// TwinCAT 3 PLC project PLC1
// ProgramVersion: 3.1.4024.0
// libraries:
//   Tc2_MC2, * (Beckhoff Automation GmbH)
//   Tc2_Standard, * (Beckhoff Automation GmbH)
//   Tc2_System, * (Beckhoff Automation GmbH)
//   Tc2_TcpIp, * (Beckhoff Automation GmbH)
//   Tc3_Module, * (Beckhoff Automation GmbH)
// project tree:
//   DUTs/ E_MelsecDevice.TcDUT, ST_MelsecSession.TcDUT, ST_Point2D.TcDUT, ST_QD75_Command.TcDUT, ST_QD75_Feedback.TcDUT
//   GVLs/ GVL.TcGVL
//   / PlcTask.TcTTO
//   POUs/ FB_ConveyorEncoder.TcPOU, FB_ConveyorTracking4Pt.TcPOU, FB_EziServoControl.TcPOU, FB_MelsecRead.TcPOU, FB_MelsecTcpConfig.TcPOU, FB_MelsecWrite.TcPOU, FB_QD75CommandPublisher.TcPOU, MAIN.TcPOU
// real-time tasks:
//   TASK PlcTask: cycle T#10ms, priority 20, ADS port 350
// motion (NC):
//   TASK NC-Task 1 SAF: cycle T#2ms, priority 4, ADS port 501
//   TASK NC-Task 1 SVB: cycle T#10ms, priority 8, ADS port 511
//   AXIS Axis 1 (id 2)
//     General: UnitName=Degree
//     Velo: Maximum=50000
//     OtherSettings: AllowMotionCmdToSlave=true
//     encoder EncType=19
//       EncPara: ScaleFactorNumerator=360, ScaleFactorDenominator=10000, MaxCount=#xffffffff
//     drive DrvType=16
//       DrvPara: MaxCount=#xffffffff, DriveControlDWord=#x00020000
//         Analog: VeloReferenz=60000, TorqueSetpointScale=10, ScaleFactorActTorque=0.1
//         TimeComp: TaskDelayCycles=1
//     controller CtrType=1
//       CtrPara: PriorControlFactor=1
//         PosDiffControl: Range=60, Time=0.05
//         Observer: BandWidth=20
// I/O:
//   DEVICE Device 2 (EtherCAT), AmsNetId 10.81.27.140.3.1
//     Box 1 (NA-9286,Crevis) [NA-9286 EtherCAT Adapter, Crevis]
//       modules: Module 1 (ST-5101), Module 2 (ST-1228), Module 3 (ST-1228), Module 4 (ST-1228), Module 5 (ST-1228), Module 6 (ST-1228), Module 7 (ST-2318), Module 8 (ST-2318), Module 9 (ST-2318), Module 10 (ST-2318), Module 11 (ST-4424), Module 12 (ST-5114), Module 13 (ST-3214)
//     Drive 2 (Ezi-SERVO2 EtherCAT) [Ezi-SERVO2 EtherCAT]
// variable links:
//   NC-Task 1 SAF/Axes/Axis 1 <-> Device 2 (EtherCAT)/Drive 2 (Ezi-SERVO2 EtherCAT)
//     Drive/Inputs/In/nDcOutputTime <-> InfoData/DcOutputShift
//     Drive/Inputs/In/nState1 <-> CSP Inputs/Status Word
//     Drive/Inputs/In/nState2 <-> CSP Inputs/Status Word @bit 8
//     Drive/Inputs/In/nState4 @bit 1 <-> WcState/InputToggle
//     Drive/Inputs/In/nState4 <-> WcState/WcState
//     Drive/Outputs/Out/nCtrl1 <-> CSP Outputs/Control Word
//     Drive/Outputs/Out/nCtrl2 <-> CSP Outputs/Control Word @bit 8
//     Drive/Outputs/Out/nDataOut1 <-> CSP Outputs/Target Position
//     Enc/Inputs/In/nDataIn1 <-> CSP Inputs/Position Actual Value
//     Enc/Inputs/In/nDataIn3 <-> CSP Inputs/Touch probe 1 positive value
//     Enc/Inputs/In/nDataIn5 <-> CSP Inputs/Touch probe 2 positive value
//     Enc/Inputs/In/nDcInputTime <-> InfoData/DcInputShift
//     Enc/Inputs/In/nState4 @bit 1 <-> WcState/InputToggle
//     Enc/Inputs/In/nState4 <-> WcState/WcState
//     Enc/Inputs/In/nState5 <-> CSP Inputs/Touch probe status
//     Enc/Inputs/In/nState6 <-> CSP Inputs/Touch probe status @bit 8
//     Enc/Outputs/Out/nCtrl5 <-> CSP Outputs/Touch probe function
//     Enc/Outputs/Out/nCtrl6 <-> CSP Outputs/Touch probe function @bit 8
//   PLC1/PLC1 Instance <-> Device 2 (EtherCAT)/Box 1 (NA-9286,Crevis)
//     PlcTask Inputs/GVL.aIn[{0..15}] <-> Module 12 (ST-5114)/Input(s)/Byte {0..15}  (16 links)
//     PlcTask Outputs/GVL.aOut[{0..3}] <-> Module 12 (ST-5114)/Output(s)/Byte {0..3}  (4 links)
//   PLC1/PLC1 Instance <-> NC-Task 1 SAF/Axes/Axis 1
//     PlcTask Inputs/MAIN.Axis1.NcToPlc <-> Outputs/ToPlc
//     PlcTask Outputs/MAIN.Axis1.PlcToNc <-> Inputs/FromPlc

CONFIGURATION PLC1
    RESOURCE PLC ON TwinCAT3
        TASK PlcTask(INTERVAL := T#10ms, PRIORITY := 20);
        PROGRAM MAIN WITH PlcTask : MAIN;
    END_RESOURCE
END_CONFIGURATION

// ---- DUTs/E_MelsecDevice.TcDUT
// Mã định danh vùng nhớ phần cứng Mitsubishi theo chuẩn MC Protocol Binary 3E Frame
TYPE E_MelsecDevice :
(
    DEV_D   := 16#A8, // Thanh ghi dữ liệu D (Data Register) - Word
    DEV_M   := 16#90, // Rơ-le nội bộ M (Internal Relay) - Bit / Word
    DEV_W   := 16#B4, // Thanh ghi liên kết W (Link Register) - Word
    DEV_R   := 16#AF, // Thanh ghi tệp R (File Register) - Word
    DEV_ZR  := 16#B0, // Thanh ghi tệp liên tục ZR (File Register Consecutive) - Word
    DEV_X   := 16#9C, // Ngõ vào vật lý X (Input) - Bit
    DEV_Y   := 16#9D, // Ngõ ra vật lý Y (Output) - Bit
    DEV_B   := 16#A0, // Rơ-le liên kết B (Link Relay) - Bit / Word
    DEV_L   := 16#92, // Rơ-le chốt L (Latch Relay) - Bit
    DEV_TN  := 16#C2, // Giá trị hiện tại Timer TN (Timer Current Value) - Word
    DEV_CN  := 16#C5  // Giá trị hiện tại Counter CN (Counter Current Value) - Word
);
END_TYPE

// ---- DUTs/ST_MelsecSession.TcDUT
TYPE ST_MelsecSession :
STRUCT
    hSocket     : T_HSOCKET; // Socket TCP dùng chung
    bConnected  : BOOL;      // TRUE khi đã kết nối PLC
    bBusy       : BOOL;      // TRUE khi Read hoặc Write đang giao dịch
    bError      : BOOL;      // Lỗi cuối cùng
    nErrorID    : UDINT;     // Mã lỗi cuối cùng
END_STRUCT
END_TYPE

// ---- DUTs/ST_Point2D.TcDUT
TYPE ST_Point2D :
STRUCT
    X : LREAL; // Tọa độ X (mm)
    Y : LREAL; // Tọa độ Y (mm)
END_STRUCT
END_TYPE

// ---- DUTs/ST_QD75_Command.TcDUT
TYPE ST_QD75_Command :
STRUCT
    Target_X       : DINT; // D100..D101: Tọa độ đón đầu trục X (0.1 um)
    Target_Y       : DINT; // D102..D103: Tọa độ trục Y đỉnh (0.1 um)
    Target_Z_Down  : DINT; // D104..D105: Độ cao hạ chấm keo (0.1 um, 4.0mm = 40000)
    Speed_Approach : DINT; // D106..D107: Vận tốc bay nội suy 3 trục (0.01 mm/min, 500mm/s = 3000000)
    Speed_Sync     : DINT; // D108..D109: Vận tốc đồng tốc trục X khi chấm keo (= V_conv * 6000)
    DeltaX_Sync    : DINT; // D110..D111: Quãng đường trượt đồng tốc 60ms (0.1 um)
    Target_Z_Safe  : DINT; // D112..D113: Độ cao an toàn khi rút kim (0.1 um, 0.0mm = 0)
    Vertex_Index   : INT;  // D114: Thứ tự đỉnh đang làm (1..4)
END_STRUCT
END_TYPE

// ---- DUTs/ST_QD75_Feedback.TcDUT
TYPE ST_QD75_Feedback :
STRUCT
    Ack_Done    : BOOL; // M1001: PLC-Q báo Point 3 hoàn tất
    Robot_Busy  : BOOL; // M102: PLC-Q đang kiểm tra/nạp/chạy
    In_Position : BOOL; // M103: Đỉnh đã hoàn tất, chờ Master hạ M1000
    Robot_Alarm : BOOL; // M104: QD75 hoặc kiểm tra biên báo lỗi
END_STRUCT
END_TYPE

// ---- GVLs/GVL.TcGVL
VAR_GLOBAL
    aIn  AT %I* : ARRAY[0..15] OF BYTE;  // TxPDO 16 byte
    aOut AT %Q* : ARRAY[0..3]  OF BYTE;  // RxPDO 4 byte
END_VAR

// ---- POUs/MAIN.TcPOU
PROGRAM MAIN
VAR
    // ================================================================
    // 1. KẾT NỐI TCP VỚI CPU MITSUBISHI Q06UDEH (CỔNG 5010)
    // ================================================================
    stMelsec            : ST_MelsecSession; // Session TCP dùng chung
    fbMelsecConfig      : FB_MelsecTcpConfig;

    bTcpEnable          : BOOL := TRUE;     // Tự động kết nối và duy trì kết nối mạng
    sPlcQ_IP            : STRING(15) := '192.168.3.39'; // IP của PLC-Q
    nPlcQ_Port          : UDINT := 5010;   // Cổng Port MC Protocol 5010

    bPlcQConnected      : BOOL;             // ĐÈN BÁO: TRUE = Đã thông mạng với PLC-Q
    bPlcQError          : BOOL;
    nPlcQErrorID        : UDINT;

    // ================================================================
    // 2. TEST TRUYỀN THÔNG THỦ CÔNG SANG PLC-Q (KHI bStartGlueCycle = FALSE)
    // ================================================================
    bTest_WriteD100     : BOOL := FALSE;    // Click đúp TRUE -> Ghi nTest_D100_Val vào D100-D101
    nTest_D100_Val      : DINT := 100;      // Số 32-bit gửi thử sang D100
    bTest_WriteM1000    : BOOL := FALSE;    // Click đúp TRUE -> Ghi bit M1000
    bTest_M1000_Val     : BOOL := TRUE;     // Giá trị bit M1000 muốn ghi (TRUE=ON, FALSE=OFF)
    bTest_ReadM1001     : BOOL := FALSE;    // Click đúp TRUE -> Đọc bit M1001 từ PLC-Q
    bTest_M1001_Result  : BOOL;             // Giá trị M1001 đọc được từ PLC-Q

    // ================================================================
    // 3. ENCODER BĂNG TẢI: ST-5114 MODULE 12
    // ================================================================
    fbConveyor          : FB_ConveyorEncoder;

    nEncoderPulse       : UINT;            // Số xung Encoder hiện tại
    nEncoderDelta       : INT;             // Xung thay đổi trong 10 ms
    rConveyorSpeed      : LREAL;           // Vận tốc băng tải lọc mượt, mm/s
    rConveyorSpeedMPM   : LREAL;           // Vận tốc băng tải, m/phút
    rConveyorDist       : LREAL;           // Tổng quãng đường băng tải, mm

    // ================================================================
    // 4. EZI-SERVO: TRỤC QUAY ĐƠN VỊ DEGREE
    // ================================================================
    Axis1               : AXIS_REF;

    fbServo             : FB_EziServoControl;

    bServo_Enable       : BOOL := TRUE;     // TRUE = Servo ON / giữ cốt
    bServo_Reset        : BOOL := FALSE;    // TRUE một chu kỳ = Reset Alarm
    bServo_JogFwd       : BOOL := FALSE;    // TRUE = chạy thuận
    bServo_JogBwd       : BOOL := FALSE;    // TRUE = chạy nghịch

    rServo_Speed        : LREAL := 100.0;   // Degree/s
    rServo_Acc          : LREAL := 400.0;   // Degree/s2
    rServo_Dec          : LREAL := 400.0;   // Degree/s2

    bServo_Ready        : BOOL;             // TRUE = Servo ON
    rServo_ActPos_Deg   : LREAL;            // Góc thực tế, Degree
    rServo_ActVel_Deg_s : LREAL;            // Vận tốc thực tế, Degree/s

    // ================================================================
    // 5. TRACKING 4 ĐIỂM: CAMERA + ENCODER
    // ================================================================
    fbTracking4Pt       : FB_ConveyorTracking4Pt;

    bSystemReset        : BOOL := FALSE;    // TRUE một chu kỳ: reset mốc phần mềm về 0
    // Camera giả lập test
    bCameraTrigger      : BOOL := FALSE;    // FALSE -> TRUE: chốt sản phẩm mới
    rCameraCenterX      : LREAL := 50.0;    // Tâm phôi X, mm
    rCameraCenterY      : LREAL := 85.0;    // Tâm phôi Y, mm
    rCameraAngleDeg     : LREAL := 0.0;     // Góc phôi, Degree
    rProductLength      : LREAL := 40.0;    // mm
    rProductWidth       : LREAL := 40.0;    // mm

    // Kết quả debug Tracking
    bProductValid       : BOOL;
    nPulseAtCamera      : UINT;
    nPulseTravel        : INT;
    rPartTravel_mm      : LREAL;

    aCornerBase         : ARRAY[1..4] OF ST_Point2D;
    aCornerNow          : ARRAY[1..4] OF ST_Point2D;

    // ================================================================
    // 6. QD75 COMMAND PUBLISHER: ĐIỀU PHỐI 4 ĐỈNH SANG PLC-Q
    // ================================================================
    fbPublisher         : FB_QD75CommandPublisher;

    // Lệnh chu trình chấm keo
    bStartGlueCycle     : BOOL := FALSE;   // FALSE -> TRUE: kích chạy chu trình 4 đỉnh
    bAbortGlueCycle     : BOOL := FALSE;   // TRUE: dừng khẩn cấp (ghi M105)

    // Trạng thái giám sát chu trình
    bGlueCycleBusy      : BOOL;            // Đang chạy 4 đỉnh
    bGlueCycleDone      : BOOL;            // Hoàn tất cả 4 đỉnh
    bGlueCycleError     : BOOL;            // Báo lỗi
    nGlueCurVertex      : INT;             // Đỉnh đang thực hiện (1..4)
    nGlueErrorCode      : INT;             // Mã lỗi (501..503, 900..921)
END_VAR

// ================================================================
// 1. TCP CONFIG: Kết nối / tự reconnect đến PLC-Q
// ================================================================
fbMelsecConfig(
    bEnable     := bTcpEnable,
    sRemoteHost := sPlcQ_IP,
    nRemotePort := nPlcQ_Port,
    stSession   := stMelsec
);

// Biến trạng thái đưa ra ngoài để Online debug dễ
bPlcQConnected := stMelsec.bConnected;
bPlcQError     := stMelsec.bError;
nPlcQErrorID   := stMelsec.nErrorID;


// ================================================================
// 2. ENCODER BĂNG TẢI: ST-5114 INPUT BYTE 0 + BYTE 1
// ================================================================
fbConveyor(
    bByte0          := GVL.aIn[0],
    bByte1          := GVL.aIn[1],
    rK_mm           := 0.476475,
    rCycleTime      := 0.01,

    nRawPulse       => nEncoderPulse,
    nDeltaPulse     => nEncoderDelta,
    rSpeed_mm_s     => rConveyorSpeed,
    rSpeed_m_min    => rConveyorSpeedMPM,
    rTotalDist_mm   => rConveyorDist
);


// ================================================================
// 3. EZI-SERVO: ENABLE, RESET, JOG VÀ GIÁM SÁT
// ================================================================
fbServo(
    Axis            := Axis1,
    bEnable         := bServo_Enable,
    bResetFault     := bServo_Reset,
    bJogFwd         := bServo_JogFwd,
    bJogBwd         := bServo_JogBwd,
    rTargetVelocity := rServo_Speed,
    rAcc            := rServo_Acc,
    rDec            := rServo_Dec,

    bReady          => bServo_Ready,
    rActPos_Deg     => rServo_ActPos_Deg,
    rActVel_Deg     => rServo_ActVel_Deg_s
);

IF bServo_Reset THEN
    bServo_Reset := FALSE;
END_IF;


// ================================================================
// 4. TRACKING 4 ĐIỂM: CAMERA + ENCODER
// ================================================================
fbTracking4Pt(
    bResetSystem   := bSystemReset,
    bCameraResult  := bCameraTrigger,
    rCenterX_mm    := rCameraCenterX,
    rCenterY_mm    := rCameraCenterY,
    rAngleDeg      := rCameraAngleDeg,
    rLength_mm     := rProductLength,
    rWidth_mm      := rProductWidth,

    nEncoderNow    := nEncoderPulse,
    rMmPerPulse    := 0.476475,
    rXMaxLimit_mm  := 180.0,

    bProductValid  => bProductValid,
    nPulseAtCamera => nPulseAtCamera,
    nPulseTravel   => nPulseTravel,
    rTravel_mm     => rPartTravel_mm,
    aCornerBase    => aCornerBase,
    aCornerNow     => aCornerNow
);

IF bSystemReset THEN
    bSystemReset := FALSE;
END_IF;


// ================================================================
// 5. QD75 COMMAND PUBLISHER: ĐIỀU PHỐI 4 ĐỈNH & TEST THỦ CÔNG
// ================================================================
fbPublisher(
    stSession           := stMelsec,
    bStartCycle         := bStartGlueCycle,
    bAbortCycle         := bAbortGlueCycle,

    // Tọa độ 4 góc thời gian thực từ khối Tracking
    aCornerNow          := aCornerNow,
    rConveyorSpeed_mm_s := rConveyorSpeed,

    // Động học
    rFlyTime_s          := 0.120,
    rApproachSpeed_mm_s := 500.0,
    rSyncTime_s         := 0.060,
    rZDown_mm           := 4.0,
    rZSafe_mm           := 0.0,

    // Chế độ test thủ công (chỉ có tác dụng khi bStartGlueCycle = FALSE)
    bManualWriteD100    := bTest_WriteD100,
    nD100_ManualVal     := nTest_D100_Val,
    bManualWriteM1000   := bTest_WriteM1000,
    bM1000_ManualVal    := bTest_M1000_Val,
    bManualReadM1001    := bTest_ReadM1001,

    // Giám sát
    bBusy               => bGlueCycleBusy,
    bDone               => bGlueCycleDone,
    bError              => bGlueCycleError,
    nErrorCode          => nGlueErrorCode,
    nCurrentVertex      => nGlueCurVertex,
    bM1001_ReadBack     => bTest_M1001_Result
);

// Tự động nhả cờ kích test sau khi lệnh được nhận
IF bTest_WriteD100 AND NOT fbPublisher.bManualWriteD100 THEN
    bTest_WriteD100 := FALSE;
END_IF;

IF bTest_WriteM1000 AND NOT fbPublisher.bManualWriteM1000 THEN
    bTest_WriteM1000 := FALSE;
END_IF;

IF bTest_ReadM1001 AND NOT fbPublisher.bManualReadM1001 THEN
    bTest_ReadM1001 := FALSE;
END_IF;

END_PROGRAM

// ---- POUs/FB_MelsecTcpConfig.TcPOU
FUNCTION_BLOCK FB_MelsecTcpConfig
VAR_INPUT
    bEnable         : BOOL := TRUE;                 // TRUE = duy trì kết nối
    sRemoteHost     : STRING(15) := '192.168.3.39'; // IP PLC-Q
    nRemotePort     : UDINT := 5010;               // Port MC Protocol
END_VAR
VAR_IN_OUT
    stSession       : ST_MelsecSession;             // Session TCP dùng chung
END_VAR
VAR
    fbConnect       : FB_SocketConnect;
    fbClose         : FB_SocketClose;
    tonRetry        : TON;

    nState          : INT := 0;
    bConnectError   : BOOL;
    nConnectErrorID : UDINT;
END_VAR

// State:
// 0 = chờ reconnect
// 1 = phát cạnh mở TCP
// 2 = chờ kết quả kết nối
// 10 = đã kết nối
// 20 = đóng socket khi Disable

CASE nState OF

    0: // Chờ 2 giây trước khi thử kết nối / kết nối lại
        stSession.bConnected := FALSE;
        stSession.bBusy      := FALSE;

        IF NOT bEnable THEN
            tonRetry(IN := FALSE);
            stSession.bError := FALSE;
        ELSE
            tonRetry(IN := TRUE, PT := T#2S);

            IF tonRetry.Q THEN
                tonRetry(IN := FALSE);
                stSession.bError   := FALSE;
                stSession.nErrorID := 0;
                nState := 1;
            END_IF
        END_IF


    1: // Cạnh lên mở TCP Socket
        fbConnect(
            sSrvNetId   := '',
            sRemoteHost := sRemoteHost,
            nRemotePort := nRemotePort,
            bExecute    := TRUE,
            tTimeout    := T#3S,
            bError      => bConnectError,
            nErrId      => nConnectErrorID,
            hSocket     => stSession.hSocket
        );

        stSession.bBusy := TRUE;
        nState := 2;


    2: // Chờ FB_SocketConnect hoàn thành
        fbConnect(
            sSrvNetId   := '',
            sRemoteHost := sRemoteHost,
            nRemotePort := nRemotePort,
            bExecute    := FALSE,
            tTimeout    := T#3S,
            bError      => bConnectError,
            nErrId      => nConnectErrorID,
            hSocket     => stSession.hSocket
        );

        IF NOT fbConnect.bBusy THEN
            stSession.bBusy := FALSE;

            IF bConnectError THEN
                stSession.bError   := TRUE;
                stSession.nErrorID := nConnectErrorID;
                stSession.hSocket.handle := 0;
                nState := 0; // Chờ 2 giây, tự thử lại
            ELSE
                stSession.bConnected := TRUE;
                stSession.bError     := FALSE;
                nState := 10;
            END_IF
        END_IF


    10: // TCP đang kết nối tốt
        stSession.bConnected := TRUE;

        IF NOT bEnable THEN
            nState := 20;
        END_IF


    20: // Đóng TCP Socket khi Disable
        fbClose(
            sSrvNetId := '',
            hSocket   := stSession.hSocket,
            bExecute  := TRUE,
            tTimeout  := T#3S
        );

        nState := 21;


    21: // Chờ đóng xong
        fbClose(
            sSrvNetId := '',
            hSocket   := stSession.hSocket,
            bExecute  := FALSE,
            tTimeout  := T#3S
        );

        IF NOT fbClose.bBusy THEN
            stSession.hSocket.handle := 0;
            stSession.bConnected     := FALSE;
            stSession.bBusy          := FALSE;
            nState := 0;
        END_IF

END_CASE

END_FUNCTION_BLOCK

// ---- POUs/FB_ConveyorEncoder.TcPOU
FUNCTION_BLOCK FB_ConveyorEncoder
VAR_INPUT
    bByte0          : BYTE;             // GVL.aIn[0]
    bByte1          : BYTE;             // GVL.aIn[1]
    rK_mm           : LREAL := 0.476475;// mm / xung (D=54.6mm, 360 xung)
    rCycleTime      : LREAL := 0.01;    // 10ms
END_VAR
VAR_OUTPUT
    nRawPulse       : UINT;             // Xung tức thời
    nDeltaPulse     : INT;              // Lệch xung mỗi 10ms
    rSpeed_mm_s     : LREAL;            // VẬN TỐC LỌC MƯỢT (mm/s)
    rSpeed_m_min    : LREAL;            // Vận tốc hiển thị (m/phút)
    rTotalDist_mm   : LREAL;            // TỔNG QUÃNG ĐƯỜNG (mm)
END_VAR
VAR
    nPrev           : UINT;
    bInit           : BOOL := TRUE;
    // Bộ lọc trượt 20 chu kỳ (200ms) để triệt tiêu hoàn toàn rung lắc
    aDeltaBuf       : ARRAY[0..19] OF INT;
    nBufIdx         : INT := 0;
    nSumDelta       : INT;
    nIdx            : INT;
    rSpeed_Avg_Raw  : LREAL;
END_VAR

// 1. Ghép 2 byte thành số xung 16-bit
nRawPulse := BYTE_TO_UINT(bByte1) * 256 + BYTE_TO_UINT(bByte0);

IF bInit THEN
    nPrev := nRawPulse;
    bInit := FALSE;
END_IF

// 2. Tính số xung lệch chu kỳ 10ms (chống tràn số)
nDeltaPulse := TO_INT(TO_DINT(nRawPulse) - TO_DINT(nPrev));
nPrev       := nRawPulse;

// 3. Bộ lọc trung bình trượt 20 chu kỳ (200ms)
aDeltaBuf[nBufIdx] := nDeltaPulse;
nBufIdx := (nBufIdx + 1) MOD 20;

nSumDelta := 0;
FOR nIdx := 0 TO 19 DO
    nSumDelta := nSumDelta + aDeltaBuf[nIdx];
END_FOR;

// 4. CẮT ZERO KHI DỪNG (DEAD-BAND):
// Nếu trong 200ms không có xung nào (băng tải dừng), ép thẳng về 0.0 ngay lập tức!
IF nSumDelta = 0 THEN
    rSpeed_mm_s  := 0.0;
    rSpeed_m_min := 0.0;
ELSE
    // Tính vận tốc trung bình trong 200ms
    rSpeed_Avg_Raw := (TO_LREAL(nSumDelta) * rK_mm) / 0.2;

    // Lọc mượt nhẹ
    rSpeed_mm_s    := rSpeed_mm_s + 0.2 * (rSpeed_Avg_Raw - rSpeed_mm_s);

    // LÀM TRÒN 1 CHỮ SỐ THẬP PHÂN (Để mắt nhìn thấy số đứng yên đầm chắc, ví dụ 100.2 mm/s)
    rSpeed_mm_s    := DINT_TO_LREAL(LREAL_TO_DINT(rSpeed_mm_s * 10.0)) / 10.0;
    rSpeed_m_min   := DINT_TO_LREAL(LREAL_TO_DINT((rSpeed_mm_s * 60.0 / 1000.0) * 10.0)) / 10.0;
END_IF;

// 5. Tổng quãng đường tích lũy (chuẩn xác 100% không lọc)
rTotalDist_mm := rTotalDist_mm + (TO_LREAL(nDeltaPulse) * rK_mm);

END_FUNCTION_BLOCK

// ---- POUs/FB_EziServoControl.TcPOU
FUNCTION_BLOCK FB_EziServoControl
VAR_INPUT
    bEnable         : BOOL := TRUE;
    bResetFault     : BOOL := FALSE;
    bJogFwd         : BOOL := FALSE;
    bJogBwd         : BOOL := FALSE;
    rTargetVelocity : LREAL := 100.0;
    rAcc            : LREAL := 400.0;
    rDec            : LREAL := 400.0;
END_VAR
VAR_IN_OUT
    Axis            : AXIS_REF;
END_VAR
VAR_OUTPUT
    bReady          : BOOL;
    rActPos_Deg     : LREAL;
    rActVel_Deg     : LREAL;
END_VAR
VAR
    fbPower         : MC_Power;
    fbMoveVelocity  : MC_MoveVelocity;
    fbHalt          : MC_Halt;
    fbReset         : MC_Reset;

    rTargetVel_Prev : LREAL;
    bVelChanged     : BOOL;
    fbTrigFwd       : R_TRIG;
    fbTrigBwd       : R_TRIG;
    fbTrigStop      : R_TRIG;
END_VAR

fbReset(Axis := Axis, Execute := bResetFault);

fbPower(
    Axis            := Axis,
    Enable          := bEnable,
    Enable_Positive := TRUE,
    Enable_Negative := TRUE,
    Override        := 100.0,
    Status          => bReady
);

fbTrigFwd(CLK := bJogFwd);
fbTrigBwd(CLK := bJogBwd);
fbTrigStop(CLK := (NOT bJogFwd AND NOT bJogBwd));

IF rTargetVelocity <> rTargetVel_Prev THEN
    bVelChanged     := TRUE;
    rTargetVel_Prev := rTargetVelocity;
ELSE
    bVelChanged     := FALSE;
END_IF

fbMoveVelocity(
    Axis         := Axis,
    Execute      := (fbTrigFwd.Q OR fbTrigBwd.Q OR (bVelChanged AND (bJogFwd OR bJogBwd))),
    Velocity     := rTargetVelocity,
    Acceleration := rAcc,
    Deceleration := rDec,
    Jerk         := 10000.0,
    Direction    := SEL(bJogBwd, MC_Positive_Direction, MC_Negative_Direction)
);

fbHalt(
    Axis         := Axis,
    Execute      := fbTrigStop.Q,
    Deceleration := rDec,
    Jerk         := 10000.0
);

rActPos_Deg := Axis.NcToPlc.ActPos;
rActVel_Deg := Axis.NcToPlc.ActVelo;

END_FUNCTION_BLOCK

// ---- POUs/FB_ConveyorTracking4Pt.TcPOU
FUNCTION_BLOCK FB_ConveyorTracking4Pt
VAR_INPUT
    bResetSystem     : BOOL;
    bCameraResult    : BOOL;
    rCenterX_mm      : LREAL;
    rCenterY_mm      : LREAL;
    rAngleDeg        : LREAL;
    rLength_mm       : LREAL := 40.0;
    rWidth_mm        : LREAL := 40.0;
    nEncoderNow      : UINT;
    rMmPerPulse      : LREAL := 0.476475;
    rXMaxLimit_mm    : LREAL := 180.0;
END_VAR

VAR_OUTPUT
    bProductValid    : BOOL;
    nPulseAtCamera   : UINT;
    nPulseTravel     : INT;
    rTravel_mm       : LREAL;
    aCornerBase      : ARRAY[1..4] OF ST_Point2D;
    aCornerNow       : ARRAY[1..4] OF ST_Point2D;
END_VAR

VAR
    fbCameraEdge     : R_TRIG;
    rRad             : LREAL;
    rCosA            : LREAL;
    rSinA            : LREAL;
    rHalfLength      : LREAL;
    rHalfWidth       : LREAL;
    nIndex           : INT;
    bFirstScan       : BOOL := TRUE;
END_VAR

// Reset mốc phần mềm một lần khi PLC khởi động hoặc khi bResetSystem kích.
IF bFirstScan OR bResetSystem THEN
    bFirstScan     := FALSE;
    bProductValid  := FALSE;
    nPulseAtCamera := nEncoderNow;
    nPulseTravel   := 0;
    rTravel_mm     := 0.0;

    FOR nIndex := 1 TO 4 DO
        aCornerBase[nIndex].X := 0.0;
        aCornerBase[nIndex].Y := 0.0;
        aCornerNow[nIndex].X  := 0.0;
        aCornerNow[nIndex].Y  := 0.0;
    END_FOR;
END_IF;

fbCameraEdge(CLK := bCameraResult);

// Camera chụp: chốt encoder và tính bốn góc gốc.
IF fbCameraEdge.Q THEN
    nPulseAtCamera := nEncoderNow;
    nPulseTravel   := 0;
    rTravel_mm     := 0.0;

    rRad   := rAngleDeg * 3.141592653589793 / 180.0;
    rCosA  := COS(rRad);
    rSinA  := SIN(rRad);
    rHalfLength := rLength_mm / 2.0;
    rHalfWidth  := rWidth_mm / 2.0;

    aCornerBase[1].X := rCenterX_mm + rHalfLength * rCosA - rHalfWidth * rSinA;
    aCornerBase[1].Y := rCenterY_mm + rHalfLength * rSinA + rHalfWidth * rCosA;
    aCornerBase[2].X := rCenterX_mm - rHalfLength * rCosA - rHalfWidth * rSinA;
    aCornerBase[2].Y := rCenterY_mm - rHalfLength * rSinA + rHalfWidth * rCosA;
    aCornerBase[3].X := rCenterX_mm - rHalfLength * rCosA + rHalfWidth * rSinA;
    aCornerBase[3].Y := rCenterY_mm - rHalfLength * rSinA - rHalfWidth * rCosA;
    aCornerBase[4].X := rCenterX_mm + rHalfLength * rCosA + rHalfWidth * rSinA;
    aCornerBase[4].Y := rCenterY_mm + rHalfLength * rSinA - rHalfWidth * rCosA;

    FOR nIndex := 1 TO 4 DO
        aCornerNow[nIndex] := aCornerBase[nIndex];
    END_FOR;
    bProductValid := TRUE;
END_IF;

// Tracking thời gian thực theo encoder.
IF bProductValid THEN
    nPulseTravel := TO_INT(nEncoderNow - nPulseAtCamera);
    rTravel_mm   := TO_LREAL(nPulseTravel) * rMmPerPulse;

    FOR nIndex := 1 TO 4 DO
        aCornerNow[nIndex].X := aCornerBase[nIndex].X + rTravel_mm;
        aCornerNow[nIndex].Y := aCornerBase[nIndex].Y;
    END_FOR;

    // Hủy sản phẩm nếu toàn bộ cạnh phía sau đã vượt vùng X của Gantry.
    IF (aCornerNow[2].X > rXMaxLimit_mm) AND (aCornerNow[3].X > rXMaxLimit_mm) THEN
        bProductValid := FALSE;
        nPulseTravel  := 0;
        rTravel_mm    := 0.0;
    END_IF;
END_IF;

END_FUNCTION_BLOCK

// ---- POUs/FB_QD75CommandPublisher.TcPOU
FUNCTION_BLOCK FB_QD75CommandPublisher
VAR_INPUT
    // ================================================================
    // 1. ĐIỀU KHIỂN CHU TRÌNH TỰ ĐỘNG 4 ĐỈNH
    // ================================================================
    bStartCycle         : BOOL;             // Cạnh lên: bắt đầu chu trình 4 đỉnh
    bAbortCycle         : BOOL;             // Dừng khẩn cấp / Hủy chu trình

    // Dữ liệu từ khối Tracking & Băng tải
    aCornerNow          : ARRAY[1..4] OF ST_Point2D;
    rConveyorSpeed_mm_s : LREAL;

    // Thông số Gantry & Bù trôi
    rFlyTime_s          : LREAL := 0.120;  // Thời gian Gantry bay tiếp cận (120ms)
    rApproachSpeed_mm_s : LREAL := 500.0;  // Tốc độ bay tiếp cận (500 mm/s)
    rSyncTime_s         : LREAL := 0.060;  // Thời gian trượt đồng tốc X (60ms)
    rZDown_mm           : LREAL := 4.0;    // Độ cao Z hạ xuống chấm keo (4.0mm)
    rZSafe_mm           : LREAL := 0.0;    // Độ cao Z rút lên an toàn (0.0mm)

    // ================================================================
    // 2. CHẾ ĐỘ TEST THỦ CÔNG TRỰC TIẾP (KHI bStartCycle = FALSE)
    // ================================================================
    bManualWriteD100    : BOOL := FALSE;    // Click đúp TRUE -> Ghi số 32-bit vào D100-D101
    nD100_ManualVal     : DINT := 100;      // Giá trị 32-bit tùy ý bạn muốn ghi thử vào D100
    bManualWriteM1000   : BOOL := FALSE;    // Click đúp TRUE -> Ghi bit M1000 (ON hoặc OFF)
    bM1000_ManualVal    : BOOL := TRUE;     // TRUE = Bật M1000 ON, FALSE = Tắt M1000 OFF
    bManualReadM1001    : BOOL := FALSE;    // Click đúp TRUE -> Đọc bit M1001 từ PLC-Q về
END_VAR

VAR_IN_OUT
    stSession           : ST_MelsecSession; // Socket TCP dùng chung
END_VAR

VAR_OUTPUT
    // ================================================================
    // TRẠNG THÁI VÀ ĐẦU RA GIÁM SÁT
    // ================================================================
    stCommand           : ST_QD75_Command;  // Gói 15 words gửi sang D100..D114
    bCmdM1000           : BOOL;             // Trạng thái bit M1000
    bCmdM105            : BOOL;             // Trạng thái bit M105 (Abort)
    bBusy               : BOOL;             // Đang chạy chu trình 4 đỉnh
    bDone               : BOOL;             // Đã hoàn thành cả 4 đỉnh
    bError              : BOOL;             // Báo lỗi
    nErrorCode          : INT;              // Mã lỗi (501..503, 900..921)
    nCurrentVertex      : INT;              // Đỉnh đang thực hiện (1..4)

    rTargetX_mm         : LREAL;            // Tọa độ X đón đầu (mm)
    rTargetY_mm         : LREAL;            // Tọa độ Y (mm)
    rLead_mm            : LREAL;            // Bù trôi trong thời gian bay (mm)
    rDeltaXSync_mm      : LREAL;            // Quãng trượt đồng tốc X (mm)

    bM1001_ReadBack     : BOOL;             // Giá trị M1001 đọc được từ PLC-Q
END_VAR

VAR
    fbWrite             : FB_MelsecWrite;
    fbRead              : FB_MelsecRead;

    // Biến đệm dữ liệu truyền thông
    bM1000_Value        : BOOL;
    bM105_Value         : BOOL;
    bStatusBit          : BOOL;
    nD100_SendDINT      : DINT;

    // Tham số lệnh động
    bWriteReq           : BOOL;
    bReadReq            : BOOL;
    eWriteDevice        : E_MelsecDevice;
    nWriteAddress       : UDINT;
    nWritePoints        : UINT;
    bWriteBitMode       : BOOL;
    pWriteData          : PVOID;
    nWriteDataSize      : UDINT;

    eReadDevice         : E_MelsecDevice;
    nReadAddress        : UDINT;
    nReadPoints         : UINT;
    bReadBitMode        : BOOL;
    pReadData           : PVOID;
    nReadDataSize       : UDINT;

    nCommError          : UDINT;
    tonPoll             : TON;
    tonTimeout          : TON;
    fbStartEdge         : R_TRIG;
    nState              : INT := 0;
END_VAR

fbStartEdge(CLK := bStartCycle);

// ================================================================
// XỬ LÝ DỪNG KHẨN CẤP / ABORT
// ================================================================
IF bAbortCycle THEN
    bCmdM105   := TRUE;
    bCmdM1000  := FALSE;
    bBusy      := FALSE;
    bDone      := FALSE;
    nState     := 99;
ELSE
    bCmdM105   := FALSE;
END_IF;

// ================================================================
// MÁY TRẠNG THÁI ĐIỀU PHỐI (FSM SEQUENCER)
// ================================================================
CASE nState OF

    0: // CHỜ LỆNH (IDLE)
        bBusy := FALSE;
        bCmdM1000 := FALSE;
        nCurrentVertex := 0;

        // 1. Kích hoạt chu trình tự động 4 đỉnh
        IF fbStartEdge.Q THEN
            IF NOT stSession.bConnected THEN
                bError := TRUE;
                nErrorCode := 900; // TCP chưa kết nối
            ELSE
                bDone := FALSE;
                bError := FALSE;
                nErrorCode := 0;
                bBusy := TRUE;
                nCurrentVertex := 1; // Bắt đầu từ Đỉnh 1
                nState := 20; // Đi thẳng vào tính toán và gửi Đỉnh 1 ngay lập tức
            END_IF;

        // 2. Chế độ Test thủ công: Ghi số 32-bit vào D100-D101
        ELSIF bManualWriteD100 THEN
            IF stSession.bConnected THEN
                nD100_SendDINT := nD100_ManualVal;
                eWriteDevice   := DEV_D;
                nWriteAddress  := 100;
                nWritePoints   := 2; // 2 words = 32-bit DINT
                bWriteBitMode  := FALSE;
                pWriteData     := ADR(nD100_SendDINT);
                nWriteDataSize := 4;
                bWriteReq      := TRUE;
                nState         := 70;
            ELSE
                bManualWriteD100 := FALSE;
            END_IF;

        // 3. Chế độ Test thủ công: Ghi Bit M1000 (ON hoặc OFF)
        ELSIF bManualWriteM1000 THEN
            IF stSession.bConnected THEN
                bM1000_Value   := bM1000_ManualVal;
                eWriteDevice   := DEV_M;
                nWriteAddress  := 1000;
                nWritePoints   := 1;
                bWriteBitMode  := TRUE;
                pWriteData     := ADR(bM1000_Value);
                nWriteDataSize := SIZEOF(bM1000_Value);
                bWriteReq      := TRUE;
                nState         := 70;
            ELSE
                bManualWriteM1000 := FALSE;
            END_IF;

        // 4. Chế độ Test thủ công: Đọc Bit M1001 từ PLC-Q
        ELSIF bManualReadM1001 THEN
            IF stSession.bConnected THEN
                eReadDevice   := DEV_M;
                nReadAddress  := 1001;
                nReadPoints   := 1;
                bReadBitMode  := TRUE;
                pReadData     := ADR(bStatusBit);
                nReadDataSize := SIZEOF(bStatusBit);
                bReadReq      := TRUE;
                nState        := 80;
            ELSE
                bManualReadM1001 := FALSE;
            END_IF;
        END_IF;

    // --- CÁC BƯỚC TEST THỦ CÔNG ---
    70: // Chờ ghi thủ công xong
        bWriteReq := FALSE;
        IF fbWrite.bDone THEN
            bManualWriteD100  := FALSE;
            bManualWriteM1000 := FALSE;
            nState := 0;
        ELSIF fbWrite.bError THEN
            bManualWriteD100  := FALSE;
            bManualWriteM1000 := FALSE;
            bError := TRUE;
            nErrorCode := 910;
            nState := 0;
        END_IF;

    80: // Chờ đọc thủ công xong
        bReadReq := FALSE;
        IF fbRead.bDone THEN
            bM1001_ReadBack  := bStatusBit;
            bManualReadM1001 := FALSE;
            nState := 0;
        ELSIF fbRead.bError THEN
            bManualReadM1001 := FALSE;
            bError := TRUE;
            nErrorCode := 920;
            nState := 0;
        END_IF;

    // --- CHU TRÌNH TỰ ĐỘNG 4 ĐỈNH ---
    20: // TÍNH TOÁN ĐÓN ĐẦU ĐỈNH nCurrentVertex
        rLead_mm       := rConveyorSpeed_mm_s * rFlyTime_s;
        rDeltaXSync_mm := rConveyorSpeed_mm_s * rSyncTime_s;
        rTargetX_mm    := aCornerNow[nCurrentVertex].X + rLead_mm;
        rTargetY_mm    := aCornerNow[nCurrentVertex].Y;

        // Giới hạn an toàn Gantry (0..180mm, 0..170mm, 0..52mm)
        // Nếu tọa độ phôi đang nằm ngoài khi test, tự ép vào vùng 50mm để luôn truyền được
        IF (rTargetX_mm < 5.0) OR ((rTargetX_mm + rDeltaXSync_mm) > 175.0) THEN
            rTargetX_mm := 50.0;
        END_IF;
        IF (rTargetY_mm < 5.0) OR (rTargetY_mm > 165.0) THEN
            rTargetY_mm := 85.0;
        END_IF;

        // Đóng gói D100..D114
        stCommand.Target_X       := LREAL_TO_DINT(rTargetX_mm * 10000.0);
        stCommand.Target_Y       := LREAL_TO_DINT(rTargetY_mm * 10000.0);
        stCommand.Target_Z_Down  := LREAL_TO_DINT(rZDown_mm * 10000.0);
        stCommand.Target_Z_Safe  := LREAL_TO_DINT(rZSafe_mm * 10000.0);
        stCommand.Speed_Approach := LREAL_TO_DINT(rApproachSpeed_mm_s * 6000.0);
        stCommand.Speed_Sync     := LREAL_TO_DINT(rConveyorSpeed_mm_s * 6000.0);
        stCommand.DeltaX_Sync    := LREAL_TO_DINT(rDeltaXSync_mm * 10000.0);
        stCommand.Vertex_Index   := nCurrentVertex;

        // Chuẩn bị gửi D100..D114 (15 words)
        eWriteDevice   := DEV_D;
        nWriteAddress  := 100;
        nWritePoints   := 15;
        bWriteBitMode  := FALSE;
        pWriteData     := ADR(stCommand);
        nWriteDataSize := SIZEOF(stCommand);
        bWriteReq      := TRUE;
        nState         := 21;

    21: // Chờ ghi D100..D114 hoàn tất
        bWriteReq := FALSE;
        IF fbWrite.bDone THEN
            // Bật M1000 = ON
            bCmdM1000      := TRUE;
            bM1000_Value   := TRUE;
            eWriteDevice   := DEV_M;
            nWriteAddress  := 1000;
            nWritePoints   := 1;
            bWriteBitMode  := TRUE;
            pWriteData     := ADR(bM1000_Value);
            nWriteDataSize := SIZEOF(bM1000_Value);
            bWriteReq      := TRUE;
            nState         := 22;
        ELSIF fbWrite.bError THEN
            bError := TRUE; nErrorCode := 910; nState := 99;
        END_IF;

    22: // Chờ ghi M1000 = ON hoàn tất
        bWriteReq := FALSE;
        IF fbWrite.bDone THEN
            tonTimeout(IN := TRUE, PT := T#10S); // Đếm timeout 10s chờ PLC làm xong
            nState := 30;
        ELSIF fbWrite.bError THEN
            bError := TRUE; nErrorCode := 911; nState := 99;
        END_IF;

    30: // QUÉT ĐỌC M1001 (CHỜ PLC BÁO XONG: M1001 = ON)
        tonPoll(IN := TRUE, PT := T#20MS);
        IF tonPoll.Q THEN
            tonPoll(IN := FALSE);
            eReadDevice   := DEV_M;
            nReadAddress  := 1001;
            nReadPoints   := 1;
            bReadBitMode  := TRUE;
            pReadData     := ADR(bStatusBit);
            nReadDataSize := SIZEOF(bStatusBit);
            bReadReq      := TRUE;
            nState        := 31;
        END_IF;

        IF tonTimeout.Q THEN
            bError := TRUE; nErrorCode := 920; nState := 99; // Timeout 10s
        END_IF;

    31: // Nhận kết quả đọc M1001
        bReadReq := FALSE;
        IF fbRead.bDone THEN
            bM1001_ReadBack := bStatusBit;
            IF bStatusBit THEN
                // PLC ĐÃ XONG ĐỈNH NÀY! (M1001 = ON)
                tonTimeout(IN := FALSE);
                // Hạ M1000 = OFF
                bCmdM1000      := FALSE;
                bM1000_Value   := FALSE;
                eWriteDevice   := DEV_M;
                nWriteAddress  := 1000;
                nWritePoints   := 1;
                bWriteBitMode  := TRUE;
                pWriteData     := ADR(bM1000_Value);
                nWriteDataSize := SIZEOF(bM1000_Value);
                bWriteReq      := TRUE;
                nState         := 32;
            ELSE
                nState := 30; // Chờ tiếp
            END_IF;
        ELSIF fbRead.bError THEN
            nState := 30; // retry
        END_IF;

    32: // Chờ ghi M1000 = OFF hoàn tất
        bWriteReq := FALSE;
        IF fbWrite.bDone THEN
            tonTimeout(IN := TRUE, PT := T#5S); // Timeout 5s chờ PLC hạ M1001
            nState := 40;
        ELSIF fbWrite.bError THEN
            bError := TRUE; nErrorCode := 912; nState := 99;
        END_IF;

    40: // QUÉT ĐỌC M1001 (CHỜ PLC HẠ M1001 = OFF ĐỂ RESET BẮT TAY)
        tonPoll(IN := TRUE, PT := T#20MS);
        IF tonPoll.Q THEN
            tonPoll(IN := FALSE);
            eReadDevice   := DEV_M;
            nReadAddress  := 1001;
            nReadPoints   := 1;
            bReadBitMode  := TRUE;
            pReadData     := ADR(bStatusBit);
            nReadDataSize := SIZEOF(bStatusBit);
            bReadReq      := TRUE;
            nState        := 41;
        END_IF;

        IF tonTimeout.Q THEN
            bError := TRUE; nErrorCode := 921; nState := 99;
        END_IF;

    41: // Nhận kết quả đọc M1001
        bReadReq := FALSE;
        IF fbRead.bDone THEN
            bM1001_ReadBack := bStatusBit;
            IF NOT bStatusBit THEN
                // PLC đã hạ M1001 = OFF -> SẴN SÀNG CHO ĐỈNH TIẾP THEO!
                tonTimeout(IN := FALSE);
                IF nCurrentVertex < 4 THEN
                    nCurrentVertex := nCurrentVertex + 1; // Sang đỉnh 2, 3, 4
                    nState := 20;                         // Tính và gửi đỉnh kế tiếp ngay!
                ELSE
                    // ĐÃ XONG CẢ 4 ĐỈNH!
                    bBusy := FALSE;
                    bDone := TRUE;
                    nState := 0;
                END_IF;
            ELSE
                nState := 40; // Chờ tiếp
            END_IF;
        ELSIF fbRead.bError THEN
            nState := 40;
        END_IF;

    99: // LỖI / DỪNG
        bBusy := FALSE;
        bCmdM1000 := FALSE;
        IF NOT bStartCycle AND NOT bAbortCycle THEN
            nState := 0;
        END_IF;
END_CASE;

// ================================================================
// THỰC THI GIAO DỊCH WRITE / READ QUA MC PROTOCOL
// ================================================================
fbWrite(
    stSession  := stSession,
    bExecute   := bWriteReq,
    eDevice    := eWriteDevice,
    nStartAddr := nWriteAddress,
    nPoints    := nWritePoints,
    bBitAccess := bWriteBitMode,
    pData      := pWriteData,
    nDataSize  := nWriteDataSize,
    nErrorID   => nCommError
);

fbRead(
    stSession  := stSession,
    bExecute   := bReadReq,
    eDevice    := eReadDevice,
    nStartAddr := nReadAddress,
    nPoints    := nReadPoints,
    bBitAccess := bReadBitMode,
    pData      := pReadData,
    nDataSize  := nReadDataSize,
    nErrorID   => nCommError
);

END_FUNCTION_BLOCK

// ---- POUs/FB_MelsecWrite.TcPOU
FUNCTION_BLOCK FB_MelsecWrite
VAR_INPUT
    bExecute    : BOOL;             // Cạnh lên: Bắt đầu giao dịch Write
    eDevice     : E_MelsecDevice;   // Mã vùng nhớ (DEV_D, DEV_M, ...)
    nStartAddr  : UDINT;            // Địa chỉ bắt đầu (D100 -> 100, M1000 -> 1000)
    nPoints     : UINT;             // Số điểm ghi (Số word hoặc số bit)
    bBitAccess  : BOOL;             // TRUE: Ghi bit (M), FALSE: Ghi word (D)
    pData       : PVOID;            // Con trỏ tới vùng dữ liệu nguồn
    nDataSize   : UDINT;            // Kích thước dữ liệu nguồn (bytes)
END_VAR

VAR_IN_OUT
    stSession   : ST_MelsecSession; // Session TCP dùng chung
END_VAR

VAR_OUTPUT
    bBusy       : BOOL;
    bDone       : BOOL;
    bError      : BOOL;
    nErrorID    : UDINT;            // 0=OK, Mã lỗi Beckhoff socket hoặc EndCode Mitsubishi
END_VAR

VAR
    fbTrigger   : R_TRIG;
    fbSend      : FB_SocketSend;
    fbReceive   : FB_SocketReceive;
    tonTimeout  : TON;

    aTx         : ARRAY[0..255] OF BYTE;
    aRx         : ARRAY[0..63] OF BYTE;
    nSendLength : UDINT;
    nWriteBytes : UDINT;
    nEndCode    : UINT;

    pSrcByte    : POINTER TO BYTE;
    pSrcBit     : POINTER TO BOOL;
    nIdx        : UDINT;
    nPairIdx    : UDINT;
    bBitVal1    : BYTE;
    bBitVal2    : BYTE;

    nRequestLength : UINT;
    nState      : INT := 0;
END_VAR

fbTrigger(CLK := bExecute);

// Xóa cờ trạng thái khi bắt đầu lệnh mới
IF nState = 0 THEN
    IF fbTrigger.Q THEN
        bDone    := FALSE;
        bError   := FALSE;
        nErrorID := 0;
    END_IF;
END_IF;

// Kiểm tra điều kiện tiên quyết
IF fbTrigger.Q THEN
    IF NOT stSession.bConnected THEN
        bError   := TRUE;
        nErrorID := 16#E001; // Socket chưa kết nối
        RETURN;
    ELSIF stSession.bBusy THEN
        bError   := TRUE;
        nErrorID := 16#E002; // Kênh truyền đang bận
        RETURN;
    ELSIF (pData = 0) OR (nDataSize = 0) THEN
        bError   := TRUE;
        nErrorID := 16#E003; // Con trỏ dữ liệu không hợp lệ
        RETURN;
    ELSE
        // ============================================================
        // 1. ĐÓNG GÓI KHUNG TRUYỀN MC PROTOCOL 3E FRAME (BINARY WRITE)
        // ============================================================
        // 1.1. Subheader: 0x50 0x00 (Gửi yêu cầu không giám sát)
        aTx[0] := 16#50;
        aTx[1] := 16#00;

        // 1.2. Network No: 0x00 (Mạng cục bộ)
        aTx[2] := 16#00;

        // 1.3. PC No: 0xFF (Trạm đích trực tiếp)
        aTx[3] := 16#FF;

        // 1.4. Target Module I/O No: 0xFF 0x03 (CPU đa xử lý mặc định)
        aTx[4] := 16#FF;
        aTx[5] := 16#03;

        // 1.5. Target Module Multidrop Station No: 0x00
        aTx[6] := 16#00;

        // Bytes 7..8: Request Data Length (sẽ tính và ghi sau khi nạp payload)

        // 1.6. Monitoring Timer: 0x10 0x00 (Đơn vị 250ms -> 16 = 4 giây)
        aTx[9]  := 16#10;
        aTx[10] := 16#00;

        // 1.7. Command: 0x01 0x14 (Batch Write - Ghi hàng loạt)
        aTx[11] := 16#01;
        aTx[12] := 16#14;

        // 1.8. Subcommand: 0x0001 (Bit units) hoặc 0x0000 (Word units)
        IF bBitAccess THEN
            aTx[13] := 16#01;
            aTx[14] := 16#00;
        ELSE
            aTx[13] := 16#00;
            aTx[14] := 16#00;
        END_IF;

        // 1.9. Start Device Address (3 bytes: LSB -> MSB)
        aTx[15] := UDINT_TO_BYTE(nStartAddr AND 16#FF);
        aTx[16] := UDINT_TO_BYTE(SHR(nStartAddr, 8) AND 16#FF);
        aTx[17] := UDINT_TO_BYTE(SHR(nStartAddr, 16) AND 16#FF);

        // 1.10. Device Code (M=0x90, D=0xA8, ...)
        aTx[18] := TO_BYTE(eDevice);

        // 1.11. Number of Device Points (2 bytes: LSB -> MSB)
        aTx[19] := UINT_TO_BYTE(nPoints AND 16#FF);
        aTx[20] := UINT_TO_BYTE(SHR(nPoints, 8) AND 16#FF);

        // ============================================================
        // 1.12. NẠP DỮ LIỆU CẦN GHI (WRITE PAYLOAD)
        // ============================================================
        IF bBitAccess THEN
            // Ghi Bit: MC Protocol mã hóa 2 bit vào 1 byte (Mỗi nibble 4-bit chứa 1 bit dữ liệu 0x10 / 0x01)
            pSrcBit := pData;
            nWriteBytes := (nPoints + 1) / 2; // Số byte payload

            FOR nPairIdx := 0 TO (nWriteBytes - 1) DO
                // Bit thứ nhất (nibble cao)
                IF (nPairIdx * 2) < nPoints THEN
                    IF pSrcBit[nPairIdx * 2] THEN
                        bBitVal1 := 16#10;
                    ELSE
                        bBitVal1 := 16#00;
                    END_IF;
                ELSE
                    bBitVal1 := 16#00;
                END_IF;

                // Bit thứ hai (nibble thấp)
                IF (nPairIdx * 2 + 1) < nPoints THEN
                    IF pSrcBit[nPairIdx * 2 + 1] THEN
                        bBitVal2 := 16#01;
                    ELSE
                        bBitVal2 := 16#00;
                    END_IF;
                ELSE
                    bBitVal2 := 16#00;
                END_IF;

                aTx[21 + nPairIdx] := bBitVal1 OR bBitVal2;
            END_FOR;

        ELSE
            // Ghi Word: Sao chép trực tiếp mảng bytes (Mỗi word = 2 bytes)
            pSrcByte := pData;
            nWriteBytes := UINT_TO_UDINT(nPoints) * 2;

            IF nWriteBytes > nDataSize THEN
                nWriteBytes := nDataSize; // Chống tràn bộ đệm
            END_IF;

            FOR nIdx := 0 TO (nWriteBytes - 1) DO
                aTx[21 + nIdx] := pSrcByte[nIdx];
            END_FOR;
        END_IF;

        // 1.13. Tính Request Data Length (Từ Monitoring Timer tới hết Payload)
        // Timer(2) + Cmd(2) + Subcmd(2) + Addr(3) + Dev(1) + Points(2) + Payload = 12 + nWriteBytes
        nRequestLength := 12 + UDINT_TO_UINT(nWriteBytes);
        aTx[7] := UINT_TO_BYTE(nRequestLength AND 16#FF);
        aTx[8] := UINT_TO_BYTE(SHR(nRequestLength, 8) AND 16#FF);

        // Tổng chiều dài khung gửi đi: Subheader(2) + Net(1) + PC(1) + IO(2) + Drop(1) + Len(2) + RequestLength
        nSendLength := 9 + nRequestLength;

        bBusy  := TRUE;
        nState := 10;
    END_IF;
END_IF;


// ================================================================
// MÁY TRẠNG THÁI GIAO TIẾP SOCKET
// ================================================================
CASE nState OF

    10: // Phát lệnh gửi dữ liệu qua TCP
        fbSend(
            sSrvNetId := '',
            hSocket   := stSession.hSocket,
            cbLen     := nSendLength,
            pSrc      := ADR(aTx),
            bExecute  := TRUE,
            tTimeout  := T#3S
        );

        nState := 11;


    11: // Chờ gửi xong
        fbSend(
            sSrvNetId := '',
            hSocket   := stSession.hSocket,
            cbLen     := nSendLength,
            pSrc      := ADR(aTx),
            bExecute  := FALSE,
            tTimeout  := T#3S
        );

        IF NOT fbSend.bBusy THEN
            IF fbSend.bError THEN
                bError   := TRUE;
                nErrorID := fbSend.nErrId;
                bBusy    := FALSE;
                nState   := 0;
            ELSE
                tonTimeout(IN := TRUE, PT := T#2S);
                nState := 20;
            END_IF;
        END_IF;


    20: // Phát lệnh nhận phản hồi PLC
        fbReceive(
            sSrvNetId := '',
            hSocket   := stSession.hSocket,
            cbLen     := SIZEOF(aRx),
            pDest     := ADR(aRx),
            bExecute  := TRUE,
            tTimeout  := T#3S
        );

        nState := 21;


    21: // Chờ nhận phản hồi (Polled receive với timeout 2 giây)
        tonTimeout(IN := TRUE);
        fbReceive(
            sSrvNetId := '',
            hSocket   := stSession.hSocket,
            cbLen     := SIZEOF(aRx),
            pDest     := ADR(aRx),
            bExecute  := FALSE,
            tTimeout  := T#3S
        );

        IF NOT fbReceive.bBusy THEN
            IF fbReceive.bError THEN
                tonTimeout(IN := FALSE);
                bError   := TRUE;
                nErrorID := fbReceive.nErrId;
                bBusy    := FALSE;
                nState   := 0;

            ELSIF fbReceive.nRecBytes > 0 THEN
                // Đã nhận được dữ liệu phản hồi!
                tonTimeout(IN := FALSE);

                IF fbReceive.nRecBytes < 11 THEN
                    bError   := TRUE;
                    nErrorID := 16#E006; // Frame phản hồi quá ngắn

                ELSIF (aRx[0] <> 16#D0) OR (aRx[1] <> 16#00) THEN
                    bError   := TRUE;
                    nErrorID := 16#E007; // Sai response subheader

                ELSE
                    // End code tại byte 9..10
                    nEndCode := BYTE_TO_UINT(aRx[9]) +
                                 BYTE_TO_UINT(aRx[10]) * 256;

                    IF nEndCode = 0 THEN
                        bDone := TRUE;
                    ELSE
                        bError   := TRUE;
                        nErrorID := nEndCode; // Mã lỗi Mitsubishi
                    END_IF;
                END_IF;

                bBusy  := FALSE;
                nState := 0;

            ELSIF tonTimeout.Q THEN
                // Quá 2 giây không có phản hồi
                tonTimeout(IN := FALSE);
                bError   := TRUE;
                nErrorID := 16#E008; // Timeout chờ response PLC
                bBusy    := FALSE;
                nState   := 0;

            ELSE
                // Chưa có dữ liệu về trong scan này -> Kích đọc tiếp ở scan sau
                nState := 20;
            END_IF;
        END_IF;

END_CASE;

// Cập nhật trạng thái bận vào session dùng chung
stSession.bBusy := bBusy;

END_FUNCTION_BLOCK

// ---- POUs/FB_MelsecRead.TcPOU
FUNCTION_BLOCK FB_MelsecRead
VAR_INPUT
    bExecute    : BOOL;             // Cạnh lên: Bắt đầu giao dịch Read
    eDevice     : E_MelsecDevice;   // Loại vùng nhớ (DEV_M, DEV_D, ...)
    nStartAddr  : UDINT;            // Địa chỉ bắt đầu (M1001 -> 1001, D100 -> 100)
    nPoints     : UINT;             // Số điểm đọc (Số bit hoặc số word)
    bBitAccess  : BOOL;             // TRUE: Đọc Bit (M), FALSE: Đọc Word (D)
    pData       : PVOID;            // Con trỏ tới vùng đệm lưu kết quả đọc
    nDataSize   : UDINT;            // Kích thước vùng đệm đích (bytes)
END_VAR

VAR_IN_OUT
    stSession   : ST_MelsecSession; // Session TCP dùng chung
END_VAR

VAR_OUTPUT
    bBusy       : BOOL;
    bDone       : BOOL;
    bError      : BOOL;
    nErrorID    : UDINT;            // 0=OK, Mã lỗi Beckhoff socket hoặc EndCode Mitsubishi
END_VAR

VAR
    fbTrigger   : R_TRIG;
    fbSend      : FB_SocketSend;
    fbReceive   : FB_SocketReceive;
    tonTimeout  : TON;

    aTx         : ARRAY[0..31] OF BYTE;
    aRx         : ARRAY[0..255] OF BYTE;
    nEndCode    : UINT;

    pDestByte   : POINTER TO BYTE;
    pDestBit    : POINTER TO BOOL;
    nIdx        : UDINT;
    nCopyBytes  : UDINT;

    nState      : INT := 0;
END_VAR

fbTrigger(CLK := bExecute);

// Xóa cờ trạng thái khi bắt đầu lệnh mới
IF nState = 0 THEN
    IF fbTrigger.Q THEN
        bDone    := FALSE;
        bError   := FALSE;
        nErrorID := 0;
    END_IF;
END_IF;

// Kiểm tra điều kiện tiên quyết
IF fbTrigger.Q THEN
    IF NOT stSession.bConnected THEN
        bError   := TRUE;
        nErrorID := 16#E101; // Socket chưa kết nối
        RETURN;
    ELSIF stSession.bBusy THEN
        bError   := TRUE;
        nErrorID := 16#E102; // Session đang bận
        RETURN;
    ELSIF (pData = 0) OR (nDataSize = 0) THEN
        bError   := TRUE;
        nErrorID := 16#E103; // Vùng đệm đích không hợp lệ
        RETURN;
    ELSE
        // ============================================================
        // 1. ĐÓNG GÓI KHUNG YÊU CẦU ĐỌC MC PROTOCOL 3E (BINARY READ)
        // Chiều dài cố định: 21 bytes
        // ============================================================
        // 1.1. Subheader: 0x50 0x00
        aTx[0] := 16#50;
        aTx[1] := 16#00;

        // 1.2. Network No: 0x00
        aTx[2] := 16#00;

        // 1.3. PC No: 0xFF
        aTx[3] := 16#FF;

        // 1.4. Target Module I/O: 0xFF 0x03
        aTx[4] := 16#FF;
        aTx[5] := 16#03;

        // 1.5. Target Module Drop: 0x00
        aTx[6] := 16#00;

        // 1.6. Request Data Length: 12 bytes (Từ Timer đến hết Points: 2+2+2+3+1+2 = 12)
        aTx[7] := 16#0C;
        aTx[8] := 16#00;

        // 1.7. Monitoring Timer: 0x10 0x00 (4 giây)
        aTx[9]  := 16#10;
        aTx[10] := 16#00;

        // 1.8. Command: 0x01 0x04 (Batch Read - Đọc hàng loạt)
        aTx[11] := 16#01;
        aTx[12] := 16#04;

        // 1.9. Subcommand: 0x0001 (Bit units) hoặc 0x0000 (Word units)
        IF bBitAccess THEN
            aTx[13] := 16#01;
            aTx[14] := 16#00;
        ELSE
            aTx[13] := 16#00;
            aTx[14] := 16#00;
        END_IF;

        // 1.10. Start Device Address (3 bytes: LSB -> MSB)
        aTx[15] := UDINT_TO_BYTE(nStartAddr AND 16#FF);
        aTx[16] := UDINT_TO_BYTE(SHR(nStartAddr, 8) AND 16#FF);
        aTx[17] := UDINT_TO_BYTE(SHR(nStartAddr, 16) AND 16#FF);

        // 1.11. Device Code (M=0x90, D=0xA8, ...)
        aTx[18] := TO_BYTE(eDevice);

        // 1.12. Number of Device Points (2 bytes: LSB -> MSB)
        aTx[19] := UINT_TO_BYTE(nPoints AND 16#FF);
        aTx[20] := UINT_TO_BYTE(SHR(nPoints, 8) AND 16#FF);

        bBusy  := TRUE;
        nState := 10;
    END_IF;
END_IF;


// ================================================================
// MÁY TRẠNG THÁI GIAO TIẾP SOCKET
// ================================================================
CASE nState OF

    10: // PHÁT LỆNH GỬI KHUNG REQUEST
        fbSend(
            sSrvNetId := '',
            hSocket   := stSession.hSocket,
            cbLen     := 21,
            pSrc      := ADR(aTx),
            bExecute  := TRUE,
            tTimeout  := T#3S
        );

        nState := 11;


    11: // CHỜ GỬI XONG
        fbSend(
            sSrvNetId := '',
            hSocket   := stSession.hSocket,
            cbLen     := 21,
            pSrc      := ADR(aTx),
            bExecute  := FALSE,
            tTimeout  := T#3S
        );

        IF NOT fbSend.bBusy THEN
            IF fbSend.bError THEN
                bError   := TRUE;
                nErrorID := fbSend.nErrId;
                bBusy    := FALSE;
                nState   := 0;
            ELSE
                tonTimeout(IN := TRUE, PT := T#2S);
                nState := 20;
            END_IF;
        END_IF;


    20: // PHÁT LỆNH NHẬN RESPONSE
        fbReceive(
            sSrvNetId := '',
            hSocket   := stSession.hSocket,
            cbLen     := SIZEOF(aRx),
            pDest     := ADR(aRx),
            bExecute  := TRUE,
            tTimeout  := T#3S
        );

        nState := 21;


    21: // CHỜ PLC-Q TRẢ RESPONSE (Polled receive với timeout 2 giây)
        tonTimeout(IN := TRUE);
        fbReceive(
            sSrvNetId := '',
            hSocket   := stSession.hSocket,
            cbLen     := SIZEOF(aRx),
            pDest     := ADR(aRx),
            bExecute  := FALSE,
            tTimeout  := T#3S
        );

        IF NOT fbReceive.bBusy THEN
            IF fbReceive.bError THEN
                tonTimeout(IN := FALSE);
                bError   := TRUE;
                nErrorID := fbReceive.nErrId;
                bBusy    := FALSE;
                nState   := 0;

            ELSIF fbReceive.nRecBytes > 0 THEN
                // Đã nhận được dữ liệu phản hồi!
                tonTimeout(IN := FALSE);

                IF fbReceive.nRecBytes < 11 THEN
                    bError   := TRUE;
                    nErrorID := 16#E104; // Response ngắn hơn frame tối thiểu

                ELSIF (aRx[0] <> 16#D0) OR (aRx[1] <> 16#00) THEN
                    bError   := TRUE;
                    nErrorID := 16#E105; // Sai response header

                ELSE
                    // End Code của Mitsubishi ở byte 9 và 10
                    nEndCode := BYTE_TO_UINT(aRx[9]) +
                                 BYTE_TO_UINT(aRx[10]) * 256;

                    IF nEndCode <> 0 THEN
                        bError   := TRUE;
                        nErrorID := nEndCode;

                    ELSE
                        // Dữ liệu bắt đầu tại Byte 11 của response
                        IF bBitAccess THEN
                            // Đọc Bit: Trong MC Protocol Binary, mỗi bit trả về 1 nibble (0x10 hoặc 0x01)
                            pDestBit := pData;
                            FOR nIdx := 0 TO (nPoints - 1) DO
                                IF nIdx < nDataSize THEN
                                    IF (nIdx MOD 2) = 0 THEN
                                        // Bit chẵn nằm ở nibble cao (0x10)
                                        pDestBit[nIdx] := ((aRx[11 + (nIdx / 2)] AND 16#10) <> 0);
                                    ELSE
                                        // Bit lẻ nằm ở nibble thấp (0x01)
                                        pDestBit[nIdx] := ((aRx[11 + (nIdx / 2)] AND 16#01) <> 0);
                                    END_IF;
                                END_IF;
                            END_FOR;
                        ELSE
                            // Đọc Word: Sao chép mảng bytes từ vị trí 11 sang bộ đệm đích
                            pDestByte  := pData;
                            nCopyBytes := UINT_TO_UDINT(nPoints) * 2;
                            IF nCopyBytes > (fbReceive.nRecBytes - 11) THEN
                                nCopyBytes := fbReceive.nRecBytes - 11;
                            END_IF;
                            IF nCopyBytes > nDataSize THEN
                                nCopyBytes := nDataSize;
                            END_IF;

                            FOR nIdx := 0 TO (nCopyBytes - 1) DO
                                pDestByte[nIdx] := aRx[11 + nIdx];
                            END_FOR;
                        END_IF;

                        bDone := TRUE;
                    END_IF;
                END_IF;

                bBusy  := FALSE;
                nState := 0;

            ELSIF tonTimeout.Q THEN
                // Quá 2 giây không có phản hồi
                tonTimeout(IN := FALSE);
                bError   := TRUE;
                nErrorID := 16#E103; // Timeout chờ response
                bBusy    := FALSE;
                nState   := 0;

            ELSE
                // Chưa có dữ liệu về trong scan này -> Kích đọc tiếp ở scan sau
                nState := 20;
            END_IF;
        END_IF;

END_CASE;

// Cập nhật trạng thái bận vào session dùng chung
stSession.bBusy := bBusy;

END_FUNCTION_BLOCK
